DATA_BLOCK "GDB_ConfigSetTest"
{ S7_Optimized_Access := 'TRUE' }
VERSION : 0.1
NON_RETAIN
VAR
    Corrupt : Bool;
    SetName : String[80];
    Field : Int;
    Text : String[80];
    Slot {ExternalWritable := 'False'} : Int;
    RecordScope {ExternalWritable := 'False'} : String[80];
    RecordKey {ExternalWritable := 'False'} : String[160];
END_VAR
BEGIN
END_DATA_BLOCK
